(* IEC 61131-3 sources: repolevel_ST_code_completion/extract_code/重型运输系统/core/struct, 11 files *)

(* ---- CmdPercentSet.st ---- *)
TYPE CmdPercentSet :
STRUCT
	extendPercent		:WORD;		//0-65535
	retractPercent		:WORD;		//0-65535
END_STRUCT
END_TYPE

(* ---- DeviceUnit.st ---- *)
TYPE DeviceUnit :
STRUCT

	sensor			:SensorInfo;		//传感器参数
	ctrl			:DevPid;			//pid等计算控制执行参数

	vector			:TargetDirect;		//指令运行方向 1-伸出 2-缩回 3-停止
	state			:DevStatus;			//设备状态 0-未知 1-运行 2-伸出到位 3-缩回到位 4-错误

	timeCounter		:INT;				//timeoutCounter超时计数器
	exeCounter		:INT;				//ExecuteCounter额外执行时间计数

	current			:ARRAY[1..2] OF WORD;	//电流mA	[i,j] -> 地轨挡板i的电流，j=1伸出电流，j=2缩回电流

END_STRUCT
END_TYPE

(* ---- DevPid.st ---- *)
TYPE DevPid :
STRUCT
	pos			:PidParam;			//位置pid参数
	spd			:PidParam;			//速度pid参数
	ff			:FeedForward;		//前馈参数
//	dp			:DynamicPlanning;	//规划参数
	exPct		:REAL;				//伸出默认比例量0-100
	rtPct		:REAL;				//缩回默认比例量0-100

	isError		:BOOL;				//当传感器数据为0时，报错并不执行pid

	extVal		:REAL;				//设定伸出位移值
	rtcVal		:REAL;				//设定缩回位移值

END_STRUCT
END_TYPE

(* ---- DevStatus.st ---- *)
{attribute 'qualified_only'}
{attribute 'strict'}
TYPE DevStatus :
(
	unknown 	:= 0,

	runing		:= 1,

	extended	:= 2,

	retracted	:= 3,

	error		:= 4
);
END_TYPE

(* ---- FeedForward.st ---- *)
TYPE FeedForward :
STRUCT

	pstThreshold	:REAL;	//正向设定阈值
	pstKv			:REAL;
	pstKa			:REAL;
	pstKaa			:REAL;
	negThreshold	:REAL;	//反向设定阈值
	negKv			:REAL;
	negKa			:REAL;
	negKaa			:REAL;

//	pstFactor		:REAL;	//正向设定速度系数因子
//	negFactor		:REAL;	//反向设定速度系数因子

END_STRUCT
END_TYPE

(* ---- PidParam.st ---- *)
TYPE PidParam :
STRUCT
	Kp			:REAL;
	Ki			:REAL;
	Kd			:REAL;
	Set_Point	:REAL;
	Max_Val		:REAL;
	Max_ACC		:REAL;
	Act_Val		:REAL;
	Err			:REAL;
	OUT			:REAL;
END_STRUCT
END_TYPE

(* ---- SensorInfo.st ---- *)
TYPE SensorInfo :
STRUCT

	position	:REAL;	//实时位移
	speed		:REAL;	//实时速度

	//记录最大最小位移值
	retractVal	:REAL;	//缩回到位值
	extendVal	:REAL;	//伸出到位值

END_STRUCT
END_TYPE

(* ---- TargetDirect.st ---- *)
{attribute 'qualified_only'}
{attribute 'strict'}
TYPE TargetDirect :
(
	extend 	:= 1,	//伸出

	retract := 2,	//缩回

	stop	:= 3	//停止
);
END_TYPE

(* ---- UIMode.st ---- *)
TYPE UIMode :
STRUCT
	manualButtonSet			:BOOL;		//手动复位按钮模式
	usePID					:BOOL;		//使用pid
	autoEnable				:BOOL;		//自动使能
	manualPercentSet		:BOOL;		//手动设定比例量
	manualSetPid			:BOOL;		//手动调节pid参数，可通过pid测试界面设定目标位移值

	syncExt					:BOOL;		//同步伸
	syncRct					:BOOL;		//同步缩

	hydPowerOn				:BOOL;		//液压站开启 modbus 使用
	hydPowerOff				:BOOL;		//液压站关闭 modbus 使用
	hydPowerReset			:BOOL;
END_STRUCT
END_TYPE

(* ---- UiPid.st ---- *)
TYPE UiPid :
STRUCT
	pos				:PidParam;			//位置pid参数
	spd				:PidParam;			//速度pid参数
	ff				:FeedForward;		//前馈参数

	level			:INT;				//1->地轨	2->天轨
	idx				:INT;				//挡板索引编号

	devSetPos		:REAL;				//设备中的设定位置点(用于观测)
	executeVal		:REAL;				//执行值(-100.0~+100.0)

	posBtn			:BOOL;			//位置控制按钮，按下实时更新交互参数
	rstPidBtn		:BOOL;			//reset pid param button重置pid参数按钮
	pwrPercent		:REAL;			//比例阀百分比 power-percent 0-100

	extendBtn		:BOOL;
	retractBtn		:BOOL;
	stopBtn			:BOOL;

(*	posErr			:REAL;
	posOut			:REAL;
	spdErr			:REAL;
	spdOut			:REAL;*)
END_STRUCT
END_TYPE

(* ---- UIUnit.st ---- *)
TYPE UIUnit :
STRUCT
	//cmd
	pwrEnable			:BOOL;		//比例阀使能   power-enable
	pwrPercent			:REAL;		//比例阀百分比 power-percent 0-100

	//button
	btnExtend			:BOOL;
	btnRetract			:BOOL;
	btnStop				:BOOL;
	btnLast				:TargetDirect;	//上次动作方向

	//info display
	name				:STRING;	//挡板名
	wname				:WSTRING;	//山河命名
	hzname				:WSTRING;	//hua zhong ming ming
	postion				:REAL;		//位移值
	speed				:REAL;
	extendPercent		:REAL;		//伸出百分比 extend-percent

END_STRUCT
END_TYPE
